// TIA Portal project "Projet1" (V15.1)

(* hardware
DEVICE "Station S7-1200_1"  S7-1200 Station
   slot 0: "Châssis_0"  S7-1200 Rack  Rack  V1.0
   slot 1: "PLC_1"  CPU 1215C DC/DC/DC  6ES7 215-1AG40-0XB0  V4.2
   slot 2: "SM 1278_1"  4SI IO link  6ES7 278-4BD32-0XB0  V2.1
*)

// ===== PLC "PLC_1"  CPU 1215C DC/DC/DC =====

VAR_GLOBAL   // PLC tag table "Table de variables standard"
   "Détection_roue_verte" AT %I8.0 : Bool;
   "Tag_2" AT %Q0.0 : Bool;
   "Axe_1_Sens" AT %Q0.1 : Bool;
   "Départ_cycle" AT %M0.0 : Bool;
   "Aller" AT %M0.1 : Bool;
   "Tag_5" AT %M0.3 : Bool;
   "Tag_6" AT %M0.4 : Bool;
   "Retour" AT %M0.2 : Bool;
   "Cycle_en_cours" AT %M0.5 : Bool;
   "Memoire_pour_T1" AT %M1.0 : Bool;
   "Detection_roue_NodeRed" AT %M2.0 : Bool;
   "Roue_triée" AT %M3.0 : Bool;
END_VAR

// folder: System blocks/Program resources

DATA_BLOCK "IEC_Timer_0_DB"   // DB3
{ S7_Optimized_Access := 'TRUE' }
AUTHOR : Simatic
FAMILY : IEC
NAME : IEC_TMR
VERSION : 1.0
// stored: InstanceOfName IEC_TIMER
"IEC_TIMER"
BEGIN
END_DATA_BLOCK

DATA_BLOCK "IEC_Timer_0_DB_1"   // DB4
{ S7_Optimized_Access := 'TRUE' }
AUTHOR : Simatic
FAMILY : IEC
NAME : IEC_TMR
VERSION : 1.0
// stored: InstanceOfName IEC_TIMER
"IEC_TIMER"
BEGIN
END_DATA_BLOCK

DATA_BLOCK "IEC_Timer_0_DB_2"   // DB7
{ S7_Optimized_Access := 'TRUE' }
AUTHOR : Simatic
FAMILY : IEC
NAME : IEC_TMR
VERSION : 1.0
// stored: InstanceOfName IEC_TIMER
"IEC_TIMER"
BEGIN
END_DATA_BLOCK

// folder: (top level)

DATA_BLOCK "Axe_1"   // DB1, Motion_DB
{ S7_Optimized_Access := 'TRUE' }
AUTHOR : SIMATIC
FAMILY : BasicMC
NAME : TO_PosAx
VERSION : 6.0
// stored: InstanceOfName TO_PositioningAxis
"TO_PositioningAxis"
BEGIN
   // Axis.OnlinePtoModeCU = 16#0000_0002
   // Axis.DirectionOutputEnabledCU = TRUE
   // Axis.SelectedChannel2EnumCU = %Q0.1
   // Axis.SelectedChannel1EnumCU = %Q0.0
   // Pulse.MinDeltaDeltaFrequencyCU = 0.004
   // Pulse.MaxDeltaDeltaFrequencyCU = 1.0E+10
   // Pulse.MinDeltaFrequencyCU = 0.005
   // Pulse.MaxDeltaFrequencyCU = 9.5E+9
   // Pulse.MinFrequencyCU = 1.0
   // Pulse.MaxFrequencyCU = 100000.0
   // Pulse.OutputSourceCU = 16#0000_0000
   // Axis.SelectPTO = 0
   // Axis.LengthUnit.LastDistance = -1
END_DATA_BLOCK

ORGANIZATION_BLOCK "Main"   // OB1, LAD, ProgramCycle
TITLE = "Main Program Sweep (Cycle)"
{ S7_Optimized_Access := 'TRUE' }
VERSION : 0.1
   VAR_TEMP   // added for the SCL form of the ladder/FBD networks
      _w1 : Bool;
   END_VAR
BEGIN

REGION Network 1
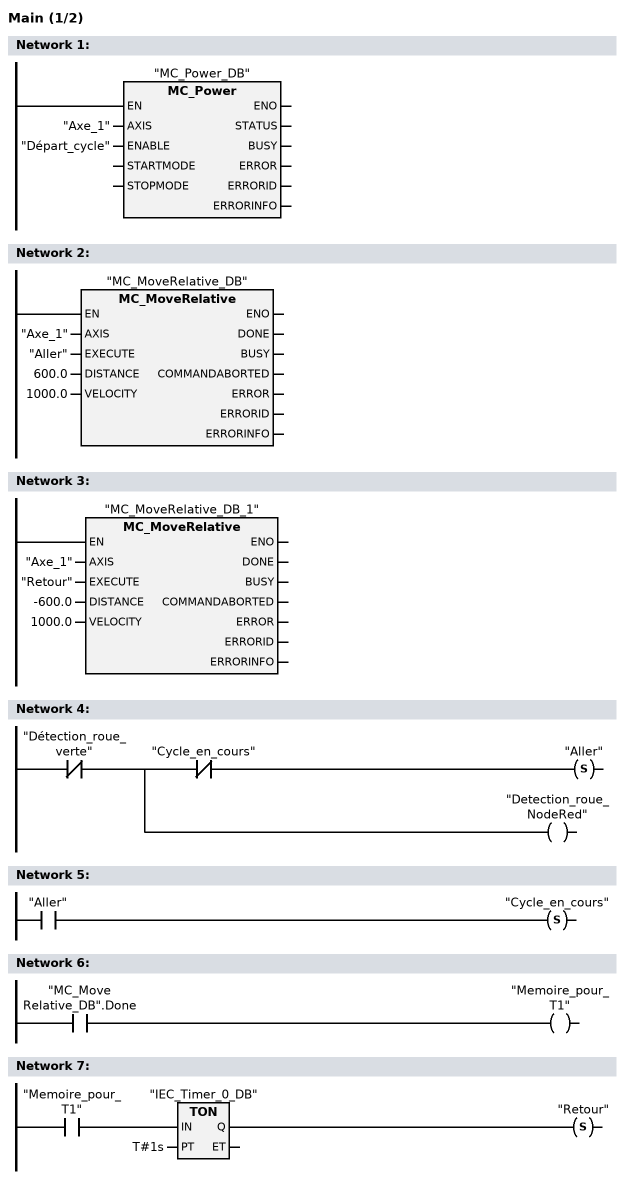
   "MC_Power_DB"(Axis := "Axe_1", Enable := "Départ_cycle");   // MC_Power
END_REGION

REGION Network 2
   "MC_MoveRelative_DB"(Axis := "Axe_1", Execute := "Aller", Distance := 600.0, Velocity := 1000.0);   // MC_MoveRelative
END_REGION

REGION Network 3
   "MC_MoveRelative_DB_1"(Axis := "Axe_1", Execute := "Retour", Distance := -600.0, Velocity := 1000.0);   // MC_MoveRelative
END_REGION

REGION Network 4
   RUNG wire#powerrail
      I_Contact( "Détection_roue_verte" )
      wire#w1
      I_Contact( "Cycle_en_cours" )
      S_Coil( "Aller" )
   END_RUNG
   RUNG wire#w1
      Coil( "Detection_roue_NodeRed" )
   END_RUNG
   // the same network as SCL:
   #_w1 := NOT "Détection_roue_verte";
   IF #_w1 AND NOT "Cycle_en_cours" THEN "Aller" := TRUE; END_IF;
   "Detection_roue_NodeRed" := #_w1;
END_REGION

REGION Network 5
   RUNG wire#powerrail
      Contact( "Aller" )
      S_Coil( "Cycle_en_cours" )
   END_RUNG
   // the same network as SCL:
   IF "Aller" THEN "Cycle_en_cours" := TRUE; END_IF;
END_REGION

REGION Network 6
   RUNG wire#powerrail
      Contact( "MC_MoveRelative_DB".Done )
      Coil( "Memoire_pour_T1" )
   END_RUNG
   // the same network as SCL:
   "Memoire_pour_T1" := "MC_MoveRelative_DB".Done;
END_REGION

REGION Network 7
   "IEC_Timer_0_DB".TON(IN := "Memoire_pour_T1", PT := T#1s);
   IF "IEC_Timer_0_DB".Q THEN "Retour" := TRUE; END_IF;
END_REGION

REGION Network 8
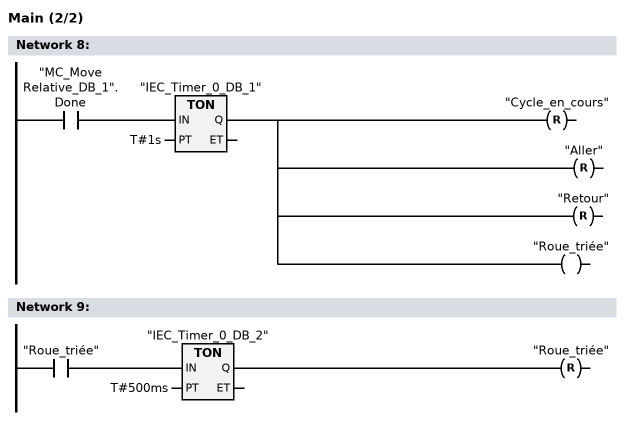
   "IEC_Timer_0_DB_1".TON(IN := "MC_MoveRelative_DB_1".Done, PT := T#1s);
   IF "IEC_Timer_0_DB_1".Q THEN
       "Cycle_en_cours" := FALSE;
       "Aller" := FALSE;
       "Retour" := FALSE;
   END_IF;
   "Roue_triée" := "IEC_Timer_0_DB_1".Q;
END_REGION

REGION Network 9
   "IEC_Timer_0_DB_2".TON(IN := "Roue_triée", PT := T#500ms);
   IF "IEC_Timer_0_DB_2".Q THEN "Roue_triée" := FALSE; END_IF;
END_REGION
END_ORGANIZATION_BLOCK